TYPE ST_ConveyorConfig :
STRUCT
    enabled : BOOL := TRUE;
    speed : LREAL := 0.75;
    startDelay : TIME := T#100ms;
END_STRUCT
END_TYPE

(* stored: Version 1.1.0.1, ProductVersion 3.1 *)
